(* IEC 61131-3 sources: PLC_Gen_Frame/Agents4PLC_release/results/task_1778475766, 1 file *)

(* ---- output.ST ---- *)
FUNCTION_BLOCK SushiConveyorControl
VAR_INPUT
    StartButton : BOOL;
    StopButton : BOOL;
    EmergencyStop : BOOL;
END_VAR
VAR_OUTPUT
    ConveyorMotor : BOOL;
END_VAR

// Generated by DummyPLCGenerator

END_FUNCTION_BLOCK
